// TIA Portal V20 export
// export: Created 2026-10-12T16:46:20.0324597Z, ExportSetting WithDefaults, DisplayName Totally Integrated Automation Portal, DisplayVersion V20 Update 6, DisplayName TIA Portal Openness, DisplayVersion V20 Update 6, DisplayName TIA Portal Version Control Interface, DisplayVersion V20 Update 6, DisplayName SINAMICS Startdrive Advanced, DisplayVersion V20 SP1 Update 2, DisplayName SINAMICS Startdrive G110M, G120, G120C, G120D, G120P, G115D, DisplayVersion V20 SP1 Update 2, DisplayName SINAMICS Startdrive G130, G150, S120, S150, SINAMICS MV, G220, S200, S210, DisplayVersion V20 SP1 Update 2, DisplayName STEP 7 Professional, DisplayVersion V20 Update 6, DisplayName STEP 7 Safety, DisplayVersion V20 Update 2, DisplayName WinCC Basic/Comfort/Advanced, DisplayVersion V20 Update 6, DisplayName WinCC Professional, DisplayVersion V20 Update 6, DisplayName WinCC Unified, DisplayVersion V20 Update 6
DATA_BLOCK "DB_IPC_to_CPU"   // DB2
{ S7_Optimized_Access := 'TRUE' }
VERSION : 0.1
// stored: AutoNumber true, DBAccessibleFromOPCUA true, DBAccessibleFromWebserver true, IsOnlyStoredInLoadMemory false, IsRetainMemResEnabled false, IsWriteProtectedInAS false, MemoryReserve 100
   VAR
      Auftrag : Array[0..9] of "UDT_Prozessroute";
      Handbetrieb : Array[1.."c_Anzahl_Bad"] of "UDT_Handbetrieb";
      Not_Halt_Reset : Bool;
      Lampentest : Bool;   // Virtuelle Tasten fuer Baeder ohne KP8 (Bad 2, 20, 47)
      Virtuelle_Tasten : Struct
         Bad_2 : Struct
            WT_Einsetzen : Array[1..3] of Bool;
            WT_Entnehmen : Array[1..3] of Bool;
         END_STRUCT;
         Bad_20 : Struct
            WT_Einsetzen : Array[1..3] of Bool;
            WT_Entnehmen : Array[1..3] of Bool;
         END_STRUCT;
         Bad_47 : Struct
            WT_Einsetzen : Array[1..3] of Bool;
            WT_Entnehmen : Array[1..3] of Bool;   // Leerlauf-Parameter pro Bad (Zustand 1: betriebsbereit halten)
         END_STRUCT;
      END_STRUCT;
   END_VAR
   VAR RETAIN
      Leerlauf : Array[1.."c_Anzahl_Bad"] of "UDT_Peripherie_Soll";   // Standby-Parameter pro Bad (Zustand 2: abgesenkt, Energie sparen)
      Standby : Array[1.."c_Anzahl_Bad"] of "UDT_Peripherie_Soll";   // Anlagenzustand: 0=undefiniert/alles aus, 1=Leerlauf, 2=Standby
   END_VAR
   VAR
      Zustand : Array[1.."c_Anzahl_Bad"] of Int;   // PT100 Offset pro Bad (vom IPC einstellbar, in Grad Celsius)
      PT100_Offset : Array[1.."c_Anzahl_Bad"] of Real;
   END_VAR
BEGIN
   PT100_Offset[7] := -4.0;
   PT100_Offset[8] := -3.8;
   PT100_Offset[12] := -4.0;
   PT100_Offset[25] := -5.8;
   PT100_Offset[36] := -3.4;
   PT100_Offset[40] := -3.2;
   PT100_Offset[46] := -3.0;
END_DATA_BLOCK
